PROGRAM main
  VAR
    Process : FB_1_Process;
    Packaging : FB_2_Packaging;
    Motion : FB_3_Motion;
    Utilities : FB_4_Utilities;
  END_VAR
  VAR_INPUT
  END_VAR
  VAR_OUTPUT
  END_VAR

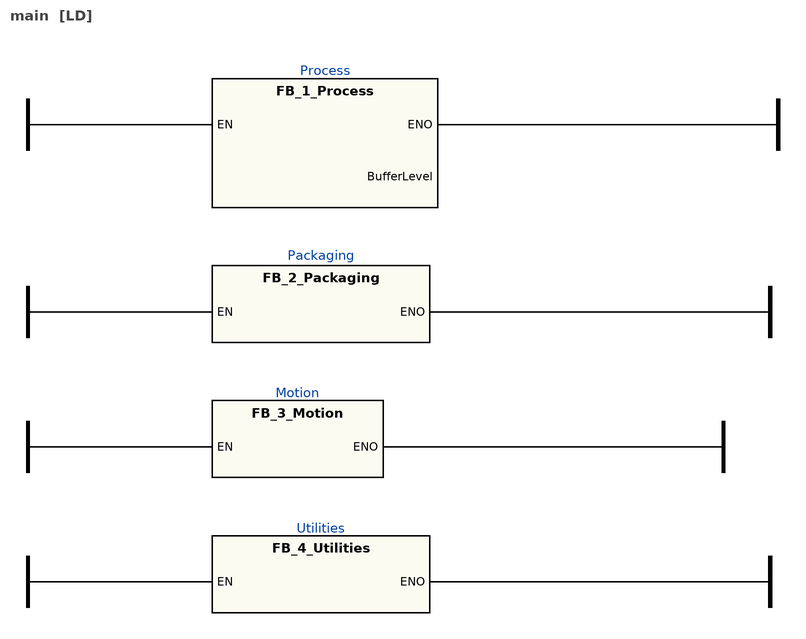
(* LD diagram, written out as Structured Text *)
Process();
Packaging();
Motion();
Utilities();
END_PROGRAM
